  rq_init_comm_if_connected(9, "1")
  rq_init_comm_if_connected(2, "2")
  rq_init_comm_if_connected(3, "3")
  rq_init_comm_if_connected(4, "4")
  rq_print_connected_grippers()
  rq_gripper_communication_thread = run rq_gripper_communication()
  set_closed_norm(97.6470588235294, 1)
  set_open_norm(1.1764705882352942, 1)
  set_closed_mm(0.0, 1)
  set_open_mm(53.0, 1)
  set_closed_norm(100.0, 2)
  set_open_norm(0.0, 2)
  set_closed_mm(0.0, 2)
  set_open_mm(50.0, 2)
  set_closed_norm(100.0, 3)
  set_open_norm(0.0, 3)
  set_closed_mm(0.0, 3)
  set_open_mm(50.0, 3)
  set_closed_norm(100.0, 4)
  set_open_norm(0.0, 4)
  set_closed_mm(0.0, 4)
  set_open_mm(50.0, 4)
  rq_current_limit_enabled = False
  while(not rq_gripper_communication_thread_started):
      sync()
  end
  # end: URCap Installation Node
  global Start_p=p[-.033064633790, -.365398531763, .389873206922, .000000000001, .000000000001, 2.725785203584]
  global Start_q=[-1.287596562866887, -1.232866726886848, -1.6880113260231102, -1.7912103151657988, 1.5729028131945846, 0.6981423183093938]
  global container_start_p=p[.200650292861, -.570238752026, .330084459991, 1.360500825815, .021700154388, 2.681649888469]
  global container_start_q=[-0.7671117850166942, -2.170180210127774, -0.8654875324671831, -2.4760661058854714, 1.019668964673781, 1.1886838746103445]
  global container_wp_1_p=p[.170613637794, -.572150573676, .294509026043, 1.259497117139, -.008270589399, 2.787717865625]
  global container_wp_1_q=[-0.8129253370121727, -2.0726598902108755, -1.0846040680899218, -2.2403146195823957, 1.0281191187839607, 1.0435744211830564]
  global Waypoint_55_p=p[.077280900603, -.567308602990, .212067617714, 1.259497117148, -.008270589399, 2.787717865619]
  global Waypoint_55_q=[-0.9181858327853867, -1.9744793804952083, -1.4540279077890048, -1.9155621911627945, 0.9643238328181578, 0.9457250675800015]
  global Waypoint_56_p=p[.135568164031, -.570867938153, .245215470413, 1.476861317558, -.018269607491, 2.679642659499]
  global Waypoint_56_q=[-0.8259784040282607, -2.108036981522602, -1.2111990877342924, -2.2405969375728745, 0.9451797152137279, 1.125710531287379]
  global Waypoint_1_p=p[.175610325005, -.574616614452, .223223522166, 1.743761338383, -.031006259154, 2.516019384206]
  global Waypoint_1_q=[-0.7669248033620333, -2.2968167722663964, -1.042289579508017, -2.484234376785108, 0.9232841478359015, 1.3091017543818342]
  global Waypoint_59_p=p[.272401132286, -.578182925380, .239561357365, 2.126997331910, .113921148153, 2.155615020515]
  global Waypoint_59_q=[-0.6600120703326624, -2.700596948663229, -0.4450863301753998, -3.1158048115172328, 0.9327830672264099, 1.686402678489685]
  global Waypoint_58_p=p[.223648508176, -.578477552733, .276546452136, 2.174288010107, -.044108754041, 2.058653287678]
  global Waypoint_58_q=[-0.7290484882560344, -2.6749849159411134, -0.44426632073579775, -3.220833992584847, 0.9665895014735898, 1.686536774549042]
  global Waypoint_60_p=p[-.013316432876, -.544772031582, .383371643081, 2.208233379808, .037543335712, 2.097559881761]
  global Waypoint_60_q=[-0.9328326161883087, -2.0999933666355775, -1.1958015693111372, -3.060905141293654, 0.690378518537611, 1.7121940951337198]
  global Waypoint_61_p=p[-.412188693372, -.356446875193, .383371643081, 1.751740964455, -.739956256289, 1.600691174920]
  global Waypoint_61_q=[-1.766185342973321, -2.0999933666355775, -1.1958015693111372, -3.060905141293654, 0.690378518537611, 1.7121940951337198]
  global Waypoint_62_p=p[-.542658707241, -.114281911009, .251261544113, 1.813043609523, -.679411528034, 1.655271622964]
  global Waypoint_62_q=[-2.158300033470912, -1.9418836862428677, -1.8142999147147894, -2.778920736683023, 0.21900622104017292, 1.8983390235012934]
  global Waypoint_63_p=p[-.549160977092, -.110180030663, .166725956353, 1.813043615357, -.679411509043, 1.655271622307]
  global Waypoint_63_q=[-2.1753688369451893, -2.0861983564907867, -1.8682963817329084, -2.6020849204097676, 0.20299747295936665, 1.9203339368361017]
  global Waypoint_68_p=p[-.333292906431, -.480744165508, .350142125738, 2.217519979286, .140864133573, 2.209123277630]
  global Waypoint_68_q=[-1.438387057796029, -1.774776476208789, -1.7081605706825291, -2.8433626113276596, 0.07508598567825443, 1.682946898281932]
  global Waypoint_3_p=p[.200650292990, -.570238752048, .330084459986, 2.169367753390, -.046205921242, 2.085892333678]
  global Waypoint_3_q=[-0.7382627064260063, -2.5628931857922193, -0.5154631582923006, -3.24517137833243, 0.9461913499132749, 1.6652139666254717]
  global Waypoint_4_p=p[.220678860874, -.585611108654, .247463403863, 2.169367753389, -.046205921242, 2.085892333680]
  global Waypoint_4_q=[-0.7354297689791203, -2.6772953387558225, -0.5042357924848311, -3.1417091800944377, 0.9493260793054743, 1.6647026060669496]
  global Waypoint_5_p=p[.116304563730, -.565093249573, .375553899018, .685157885970, .069380584882, 2.934699151616]
  global Waypoint_5_q=[-0.9554487935176637, -1.8273442988256203, -1.1597873108138153, -1.989013540482965, 1.1919078974128405, 0.7945701907431797]
  global Waypoint_6_p=p[.116304563868, -.565093249642, .339673552379, .685157837810, .069380708857, 2.934699157210]
  global Waypoint_6_q=[-0.9556225386037127, -1.8176429686669824, -1.264118303271072, -1.8944626233198951, 1.192049102037264, 0.7947821249084998]
  global Waypoint_7_p=p[.116304563814, -.565093249565, .398257664571, .685157837809, .069380708856, 2.934699157210]
  global Waypoint_7_q=[-0.9553327241572456, -1.8383075714386141, -1.0868108907169107, -2.050975816392395, 1.1917996424394106, 0.7944337598901274]
  $ 97 "Thread_1"
  thread Thread_1():
    while (True):
      $ 98 "If Start_thread≟ True "
      if (Start_thread ==   True  ):
        $ 99 "Weight_value≔get_weight()"
        global Weight_value=get_weight()
        $ 100 "Wait: 0.25"
        sleep(0.25)
        $ 101 "sync()"
        sync()
      end
    end
  end
  threadId_Thread_1 = run Thread_1()
  $ 2 "Robot Program"
  $ 3 "Script: Weight_scale_socket.script"
  def get_weight():
  	socket_open("192.168.12.190", 3002)
  	textmsg("socket opened successfully!")
  	socket_send_string("GET_WEIGHT")
  	sync()
  	sleep(0.5)
  	receiveFromServ = socket_read_ascii_float(6)
  	while (receiveFromServ[0] <1):
  		sleep(0.5)
  		receiveFromServ = socket_read_ascii_float(1)
  		textmsg("retrying read:", receiveFromServ)
  	end
  	textmsg("Received weight:", receiveFromServ[1])
  	socket_close()
  	return receiveFromServ[1]
  end
  $ 4 "Script: dosing_pid.script"
  def dosing_pid(Target_weight):
  	#kp = 0.005
  	#ki = 0.02
  	#kd = 0.2
  	#dt = 0.05
  	#current_error = 0.0
  	#Integral_error = 0.0
  	#previous_error = 0.0
  	#tilt_angle = -1.0
  	max_tilt_angle = -0.55
  	#current_pose = get_actual_tcp_pose()

  	while ( Weight_value < Target_weight and tilt_angle < max_tilt_angle):
  		Weight_value = get_weight()
  		current_error = Target_weight - Weight_value
  		Integral_error = Integral_error + current_error*dt
  		derivative = (current_error - previous_error) / dt
  		tilt_increment = (kp * current_error) + (ki * Integral_error) + (kd * derivative)
  		current_pose = get_actual_tcp_pose()
  		tilt_angle = current_pose[4]
  		new_pose = pose_trans(current_pose, p[(tilt_increment/5), 0, 0, 0, tilt_increment, 0])
  		movel(new_pose, a = 0.075, v = 0.025, t = 0, r = 0)
  		previous_error = current_error
  		sleep(dt)
  	end
  end
  $ 5 "Start_thread≔ False "
  global Start_thread=  False
  $ 6 "kp≔0.0005"
  global kp=0.0005
  $ 7 "ki≔0.002"
  global ki=0.002
  $ 8 "kd≔0.02"
  global kd=0.02
  $ 9 "dt≔0.05"
  global dt=0.05
  $ 10 "Weight_value≔get_weight()"
  global Weight_value=get_weight()
  $ 11 "Target_weight≔'Enter the Target weight to be dispensed in gm'"
  global Target_weight=request_float_from_primary_client("Enter the Target weight to be dispensed in gm")
  $ 12 "Integral_error≔0"
  global Integral_error=0
  $ 13 "current_error≔0"
  global current_error=0
  $ 14 "previous_error≔0"
  global previous_error=0
  $ 16 "tilt_angle≔-1"
  global tilt_angle=-1
  $ 17 "MoveL"
  $ 18 "Start" "breakAfter"
  movel(Start_p, a=1.2, v=0.25)
  $ 45 "Loop Weight_value<Target_weight"
  while (Weight_value<Target_weight):
    $ 46 "MoveL"
    $ 47 "container_start" "breakAfter"
    movel(container_start_p, a=0.3, v=0.1)
    $ 48 "container_wp_1" "breakAfter"
    movel(container_wp_1_p, a=0.3, v=0.05)
    $ 49 "Loop 2 times"
    Loop_2 = 0
    while (Loop_2 < 2):
      $ 50 "Waypoint_55" "breakAfter"
      global move_thread_flag_50=0
      thread move_thread_50():
        enter_critical
        move_thread_flag_50 = 1
        movel(Waypoint_55_p, a=0.5, v=0.07)
        move_thread_flag_50 = 2
        exit_critical
      end
      move_thread_flag_50 = 0
      move_thread_han_50 = run move_thread_50()
      while (True):
        local targetTcpDirection=get_target_tcp_speed()
        local stepsToRetract=tool_contact(direction=targetTcpDirection)
        if (stepsToRetract > 0):
          kill move_thread_han_50
          stopl(3.0)
          local backTrackMovement=get_actual_joint_positions_history(stepsToRetract)
          local contactPose=get_forward_kin(backTrackMovement)
          local posDir=[targetTcpDirection[0],targetTcpDirection[1],targetTcpDirection[2]]
          local retractTo=contactPose
          if (norm(posDir) > 1e-6):
            local normalizedPosDir=normalize(posDir)
            local additionalRetraction=p[normalizedPosDir[0] * -0.01, normalizedPosDir[1] * -0.01, normalizedPosDir[2] * -0.01, 0, 0, 0]
            retractTo = pose_sub(contactPose, additionalRetraction)
          end
          movel(retractTo, a=3.0, v=0.1)
          $ 51 "Until (tool_contact_detection)"
          break
        end
        sleep(1.0E-10)
        if (move_thread_flag_50 > 1):
          join move_thread_han_50
          break
        end
        sync()
      end
      $ 52 "Waypoint_56" "breakAfter"
      movel(Waypoint_56_p, a=0.3, v=0.05)
      Loop_2 = Loop_2 + 1
    end
    $ 53 "Loop 1 times"
    Loop_3 = 0
    while (Loop_3 < 1):
      $ 54 "Waypoint_1" "breakAfter"
      movel(Waypoint_1_p, a=1.2, v=0.4)
      $ 55 "Waypoint_56" "breakAfter"
      movel(Waypoint_56_p, a=0.3, v=0.05)
      Loop_3 = Loop_3 + 1
    end
    $ 56 "Waypoint_59" "breakAfter"
    movel(Waypoint_59_p, a=0.3, v=0.05)
    $ 57 "Waypoint_58" "breakAfter"
    movel(Waypoint_58_p, a=0.3, v=0.05)
    $ 58 "MoveJ"
    $ 59 "Waypoint_60" "breakAfter"
    movej(get_inverse_kin(Waypoint_60_p, qnear=Waypoint_60_q), a=0.5235987755982988, v=0.3490658503988659, r=0.05)
    $ 60 "Waypoint_61" "breakAfter"
    movej(get_inverse_kin(Waypoint_61_p, qnear=Waypoint_61_q), a=0.5235987755982988, v=0.3490658503988659, r=0.05)
    $ 61 "Waypoint_62" "breakAfter"
    movej(get_inverse_kin(Waypoint_62_p, qnear=Waypoint_62_q), a=0.5235987755982988, v=0.3490658503988659)
    $ 62 "MoveL"
    $ 63 "Waypoint_63" "breakAfter"
    movel(Waypoint_63_p, a=0.3, v=0.05)
    $ 64 "Start_thread≔ True "
    global Start_thread=  True
    $ 65 "Wait: 0.5"
    sleep(0.5)
    $ 77 "current_pose≔get_actual_tcp_pose()"
    global current_pose= get_actual_tcp_pose ()
    $ 78 "dosing_pid(Target_weight)"
    dosing_pid(Target_weight)
    $ 79 "Start_thread≔ False "
    global Start_thread=  False
    $ 81 "Weight_value≔get_weight()"
    global Weight_value=get_weight()
    $ 82 "tilt_angle≔-1"
    global tilt_angle=-1
    $ 83 "Wait: 0.5"
    sleep(0.5)
    $ 84 "MoveL"
    $ 85 "Waypoint_68" "breakAfter"
    movel(Waypoint_68_p, a=0.2, v=0.1, r=0.05)
    $ 86 "Waypoint_3" "breakAfter"
    movel(Waypoint_3_p, a=0.4, v=0.1)
    $ 87 "Integral_error≔0"
    global Integral_error=0
    $ 88 "current_error≔0"
    global current_error=0
    $ 89 "previous_error≔0"
    global previous_error=0
  end
  $ 90 "MoveL"
  $ 91 "Waypoint_4" "breakAfter"
  movel(Waypoint_4_p, a=0.4, v=0.1)
  $ 92 "Waypoint_5" "breakAfter"
  movel(Waypoint_5_p, a=0.4, v=0.06)
  $ 93 "Waypoint_6" "breakAfter"
  movel(Waypoint_6_p, a=1.2, v=0.25)
  $ 94 "Waypoint_7" "breakAfter"
  movel(Waypoint_7_p, a=1.2, v=0.25)
  $ 95 "Start" "breakAfter"
  movel(Start_p, a=0.6, v=0.15)
  $ 96 "Popup: Powder dispensed successfully..."
  popup("Powder dispensed successfully...", "Message", False, False, blocking=True)
end
